Universal Robots URScript: T006_mistralai_Devstral-Small-2-24B-Instruct-2512_edit_lazy_rep1.urscript

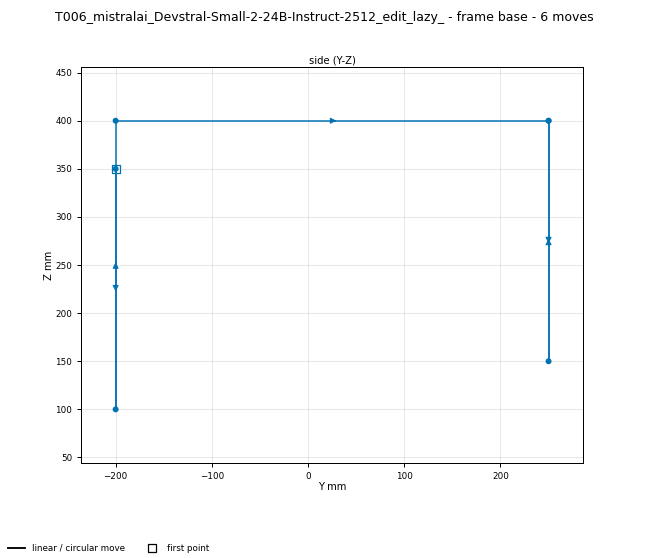
[picture p0: tool path of T006_mistralai_Devstral-Small-2-24B-Instruct-2512_edit_lazy_rep1.urscript in frame base, 6 of 8 moves have a stored position in this frame; points joined in program order, loops and branches not executed]
# Task: T006 — Bin picking with suction — fenced mode
# Improved version with optimized motion parameters and safety checks
# Operating mode: fenced | Max TCP speed: 0.400 m/s
# Robot: ur5e

def task_T006():
  # [0] Verify E-Stop clear
  if (get_digital_in(0) == True):
    popup("E-Stop active — aborting program.", error=True)
    halt
  end

  # [1] Home position
  movej([0.0000, -1.5708, 1.5708, -1.5708, -1.5708, 0.0000], a=1.4000, v=0.8750, t0=0, t1=0)

  # [2] Above bin
  movel(p[0.450000, -0.200000, 0.350000, 0.0000, 3.1416, 0.0000], a=1.5000, v=0.3500, r=0.0150, t0=0, t1=0)

  # [3] Descend into bin
  movel(p[0.450000, -0.200000, 0.100000, 0.0000, 3.1416, 0.0000], a=0.8000, v=0.1500, r=0.0150, t0=0, t1=0)

  # [4] Suction ON
  set_digital_out(0, True)

  # [5] Vacuum settle
  sleep(0.3000)

  # [6] Lift from bin
  movel(p[0.450000, -0.200000, 0.400000, 0.0000, 3.1416, 0.0000], a=1.2000, v=0.3000, r=0.0150, t0=0, t1=0)

  # [7] Transit to conveyor
  movel(p[0.450000, 0.250000, 0.400000, 0.0000, 3.1416, 0.0000], a=1.8000, v=0.3800, r=0.0200, t0=0, t1=0)

  # [8] Descend to drop
  movel(p[0.450000, 0.250000, 0.150000, 0.0000, 3.1416, 0.0000], a=1.0000, v=0.2000, r=0.0150, t0=0, t1=0)

  # [9] Suction OFF
  set_digital_out(0, False)

  # [10] Release settle
  sleep(0.2000)

  # [11] Retract above conveyor
  movel(p[0.450000, 0.250000, 0.400000, 0.0000, 3.1416, 0.0000], a=1.5000, v=0.3500, r=0.0100, t0=0, t1=0)

  # [12] Return to home
  movej([0.0000, -1.5708, 1.5708, -1.5708, -1.5708, 0.0000], a=1.4000, v=0.8750, t0=0, t1=0)

end

# Entry point
task_T006()
